# EPICS IOC start-up script: recipes-e3/iocstats/files/iocStats.iocsh
#- ### iocStats entry snippet ###
#- ####################################################
#- >> Mandatory
#- IOC - Prefix for PVs
#- ####################################################

dbLoadRecords("iocAdminSoft-ess.db", "IOC=$(IOCNAME)")
